DATA_BLOCK "GDB_LineTest"
{ S7_Optimized_Access := 'TRUE' }
VERSION : 0.1
NON_RETAIN
"FB_LineTest"
BEGIN
END_DATA_BLOCK
